FUNCTION_BLOCK TcoDriveSimpleTest EXTENDS TcoDrivesBeckhoff.TcoDriveSimple
VAR
    _serviceModeCount : ULINT;
    _serviceModeOverride : LREAL;
END_VAR
VAR
    _MC_ReadDriveAddress : MC_ReadDriveAddress;
    _fbEcCoeSdoRead : FB_EcCoeSdoRead;
    sNetId : T_AmsNetId;
    nSlaveAddr : UINT;
    _MotorType : STRING;
    _ftrig : Tc2_Standard.F_TRIG;
    _MC_ReadParameter : MC_ReadParameter;
END_VAR

SUPER^(	inEnable 			:=	inEnable,
		inEnablePositive	:=	inEnablePositive,
		inEnableNegative	:=	inEnableNegative,
		inCalibrationCam	:=	inCalibrationCam,
		inoAxisRef			:=	inoAxisRef);

END_FUNCTION_BLOCK

(* stored: Version 1.1.0.1, ProductVersion 3.1.4024.12
   POU TcoDriveSimpleTest: Id {830e1f40-136a-027f-3da2-53501fc572a7}, SpecialFunc None *)
